(* IEC 61131-3 sources: kns-port-domestic/tools/inventory_tests/fixtures/lib/src/POUs/F_Calc, 2 files *)

(* ---- F_Calc.decl.st ---- *)
// Назначение: операторы LTIME, динамическая память, запросы интерфейсов
FUNCTION F_Calc : LTIME
VAR_INPUT
    tIn : TIME;
END_VAR
VAR
    pDyn : POINTER TO INT;
    itfA : I_Base;
    itfB : I_Dev;
    udiSize : UDINT;
END_VAR

(* ---- F_Calc.impl.st ---- *)
F_Calc := TIME_TO_LTIME(tIn) + LT#1S + LTIME#2MS;
pDyn := __NEW(INT);
__DELETE(pDyn);
IF __QUERYINTERFACE(itfA, itfB) THEN
    udiSize := SIZEOF(tIn);
END_IF
{IF defined(DEBUG)}
udiSize := 0;
{END_IF}
